ABB RobotStudio station: projekt2.rspag

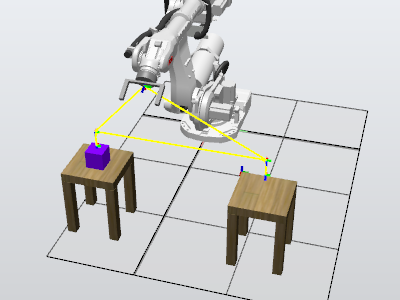
--- station ---
Station Baczyk2 (saved by RobotStudio 24.3.10958.1)
Controller Controller1
  mechanical unit ROB_1: IRB6650S_125_350_MH3_03, 6 joints, base frame (0, 0, 0) mm
Layout (positions relative to the parent item):
  - IRB6650S_125_350_MH3_03 [mechanism, from %ABB.RobotStudio.Models.IRB6650S%\IRB6650S_125_350_MH3_03.rslib] at (0, 0, 0) mm; joint values [0, 0, 0, 0, 0.5236, 0] (rad or m)
  - My_Mechanism [mechanism] at (2365.21, 0, 2010) mm, rotated rx 180 ry 60 rz 180 deg; joint values [0.16, -0.16] (rad or m)
      TCP My_Mechanism_1 at (0, 0, 90) mm
      links: L1, L2, L3
  - Group_2 [graphiccomponentgroup] at (1970.93, 882.73, 0) mm
    - Part_6 [part], size 100 x 100 x 700 mm
    - Part_7 [part], size 100 x 100 x 700 mm
    - Part_8 [part], size 100 x 100 x 700 mm
    - Part_9 [part], size 100 x 100 x 700 mm
    - Part_10 [part], size 600 x 600 x 100 mm
  - Group_3 [graphiccomponentgroup] at (1950.21, -956.94, 0) mm
    - Part_6 [part], size 100 x 100 x 700 mm
    - Part_7 [part], size 100 x 100 x 700 mm
    - Part_8 [part], size 100 x 100 x 700 mm
    - Part_9 [part], size 100 x 100 x 700 mm
    - Part_10 [part], size 600 x 600 x 100 mm
  - LineSensor_2 [smart component, from Components\LineSensor.rslib] at (2444.15, 0, 1965) mm, rotated rx 180 ry 60 rz 180 deg
      properties: Start=[0 0 0]; End=[0 0 0.15]; Length=0.15; Radius=0.01; Tag=(none); SensedPart=(none); SensedPoint=[0 0 0]
    - _sensorPart_ [part], size 20 x 20 x 150 mm
  - Attacher [smart component, from Components\Attacher.rslib]
      properties: Parent=IRB6650S_125_350_MH3_03; Flange=0; Child=(none); Mount=false; Offset=[0 0 0]; Orientation=[0 0 0]
  - Detacher [smart component, from Components\Detacher.rslib]
      properties: Child=(none); KeepPosition=true
  - Part_11 [part] at (2169.73, -741.66, 799.61) mm, size 200 x 200 x 200 mm
  - PoseMover [smart component, from Components\PoseMover.rslib]
      properties: Mechanism=My_Mechanism; Pose=1; Duration=0
  - PoseMover_2 [smart component, from Components\PoseMover.rslib]
      properties: Mechanism=My_Mechanism; Pose=2; Duration=0
  - PoseMover_3 [smart component, from Components\PoseMover.rslib]
      properties: Mechanism=My_Mechanism; Pose=1; Duration=0
Attachment: My_Mechanism is attached to IRB6650S_125_350_MH3_03 / Link6
Attachment: LineSensor_2 is attached to My_Mechanism / L2
EventTableEntry 2426: ActivationMode=2, Cyclic=false, Group=, Trigger=Gripper 2427, Actions=[EventTableActionMechanicalPose 2428], Comment=
EventTableTriggerIO 2427: Operator=0, IOValue=[1], IRC5Controller=? -1, SignalSource=Controller1 2434
EventTableActionMechanicalPose 2428: VirtualSignal=, Mechanism=My_Mechanism 2419, ToPoseName=HomePosition, VirtualSignalValue=[1]
EventTableTriggerIO 2429: Operator=0, IOValue=[0], IRC5Controller=? -1, SignalSource=Controller1 2434
EventTableEntry 2430: ActivationMode=2, Cyclic=false, Group=, Trigger=Gripper 2429, Actions=[EventTableActionMechanicalPose 2431], Comment=
EventTableActionMechanicalPose 2431: VirtualSignal=, Mechanism=My_Mechanism 2419, ToPoseName=SyncPosition, VirtualSignalValue=[1]
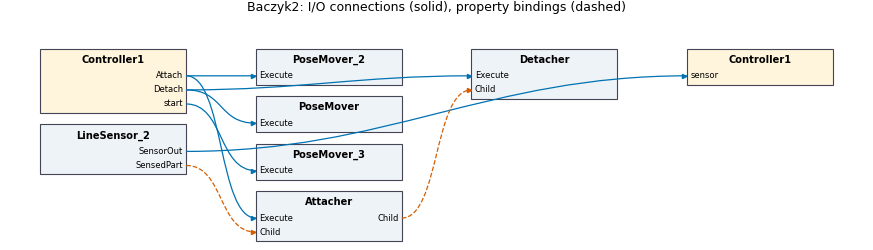
Station logic (signal -> signal, property => property):
  Controller1.Attach -> Attacher.Execute
  Controller1.Detach -> Detacher.Execute
  Controller1.Attach -> PoseMover_2.Execute
  Controller1.Detach -> PoseMover.Execute
  LineSensor_2.SensorOut -> Controller1.sensor
  Controller1.start -> PoseMover_3.Execute
  LineSensor_2.SensedPart => Attacher.Child
  Attacher.Child => Detacher.Child
Targets, tools, work objects and paths stored in the station and not in the controller backup, written as RAPID:
! task T_ROB1
MODULE Module1
  PROC Path_Flow()
    WaitTime 1;
    Set Gripper;
    WaitTime 1;
    Reset Gripper;
    WaitTime 1;
  ENDPROC
ENDMODULE


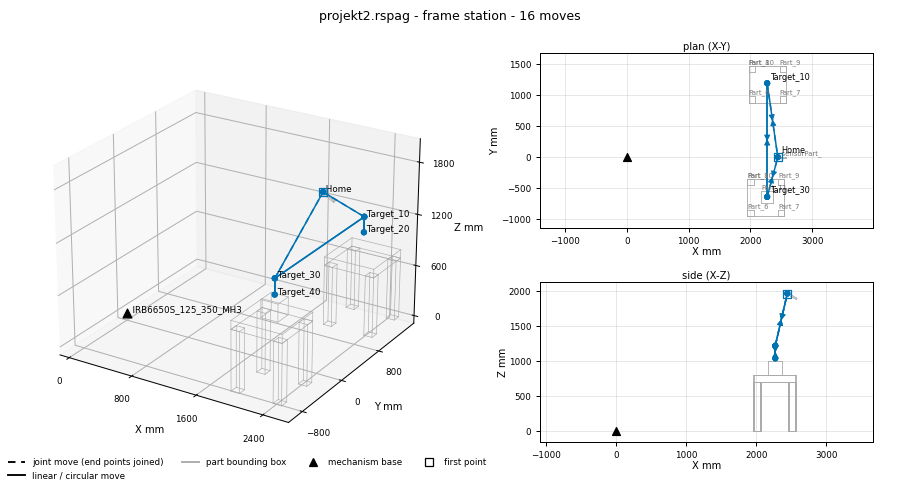
[picture p0: tool path of projekt2.rspag in frame station, 16 of 16 moves have a stored position in this frame; points joined in program order, loops and branches not executed]
--- Controller Data/Controller1/RAPID/TASK1/PROGMOD/CalibData.mod ---
MODULE CalibData
    PERS tooldata My_Mechanism_1:=[TRUE,[[0,0,90],[1,0,0,0]],[1,[0,0,90],[1,0,0,0],0,0,0]];
    TASK PERS wobjdata Workobject_2:=[FALSE,TRUE,"",[[0,0,0],[1,0,0,0]],[[0,0,0],[1,0,0,0]]];
    TASK PERS wobjdata Workobject_3:=[FALSE,TRUE,"",[[1970.926,882.727,800],[1,0,0,0]],[[0,0,0],[1,0,0,0]]];
ENDMODULE

--- Controller Data/Controller1/RAPID/TASK1/PROGMOD/Module1.mod ---
MODULE Module1
    VAR bool value;
        CONST robtarget Home:=[[472.221367097,-882.727,1165],[0.5,0,0.866025404,0],[0,0,0,0],[9E+09,9E+09,9E+09,9E+09,9E+09,9E+09]];
    CONST robtarget Target_10:=[[300.224086373,313.272936929,420.000073654],[-0.000000284,0.000000194,1,-0.000000149],[0,0,0,0],[9E+09,9E+09,9E+09,9E+09,9E+09,9E+09]];
    CONST robtarget Target_20:=[[300.224119695,313.272954476,239.999979637],[-0.000000267,0.000000194,1,-0.00000014],[0,0,0,0],[9E+09,9E+09,9E+09,9E+09,9E+09,9E+09]];
    CONST robtarget Target_30:=[[300.224073663,-1524.727216206,420.000075687],[-0.000000372,0.000000252,1,-0.00000014],[-1,-1,-1,0],[9E+09,9E+09,9E+09,9E+09,9E+09,9E+09]];
    CONST robtarget Target_40:=[[300.224095291,-1524.727007335,240.000010396],[-0.000000007,0,1,0.000000002],[-1,0,-1,0],[9E+09,9E+09,9E+09,9E+09,9E+09,9E+09]];
!***********************************************************
    !
    ! Module:  Module1
    !
    ! Description:
    !   <Insert description here>
    !
    ! Author: Mirgi
    !
    ! Version: 1.0
    !
    !***********************************************************


    !***********************************************************
    !
    ! Procedure main
    !
    !   This is the entry point of your program
    !
    !***********************************************************
    VAR bool detected;
    PROC main()
        Path_10;
    ENDPROC
    PROC Path_10()
        MoveJ Home,v1000,z100,My_Mechanism_1\WObj:=Workobject_3;
        MoveL Target_10,v1000,z100,My_Mechanism_1\WObj:=Workobject_3;
        MoveL Target_20,v1000,fine,My_Mechanism_1\WObj:=Workobject_3;
        IF sensor = 1 THEN
            PulseDO Attach;
            WaitTime 1;
            MoveL Target_10,v1000,z100,My_Mechanism_1\WObj:=Workobject_3;
            MoveL Target_30,v1000,z100,My_Mechanism_1\WObj:=Workobject_3;
            MoveL Target_40,v1000,fine,My_Mechanism_1\WObj:=Workobject_3;
            PulseDO Detach;
            WaitTime 1;
            MoveL Target_30,v1000,z100,My_Mechanism_1\WObj:=Workobject_3;
            MoveJ Home,v1000,z100,My_Mechanism_1\WObj:=Workobject_3;
        ELSE
            MoveJ Home,v1000,z100,My_Mechanism_1\WObj:=Workobject_3;
            MoveL Target_30,v1000,z100,My_Mechanism_1\WObj:=Workobject_3;
            MoveL Target_40,v1000,fine,My_Mechanism_1\WObj:=Workobject_3;
            PulseDO Attach;
            WaitTime 1;
            MoveL Target_30,v1000,z100,My_Mechanism_1\WObj:=Workobject_3;
            MoveL Target_10,v1000,z100,My_Mechanism_1\WObj:=Workobject_3;
            MoveL Target_20,v1000,fine,My_Mechanism_1\WObj:=Workobject_3;
            PulseDO Detach;
            WaitTime 1;
            MoveL Target_10,v1000,z100,My_Mechanism_1\WObj:=Workobject_3;
            MoveJ Home,v1000,z100,My_Mechanism_1\WObj:=Workobject_3;
        ENDIF
    ENDPROC
ENDMODULE

--- Controller Data/Controller1/SYSPAR/EIO.cfg ---
EIO:CFG_1.0:6:1::
#
EIO_SIGNAL:

      -Name "Gripper" -SignalType "DO" -Access "All"

      -Name "Attach" -SignalType "DO"

      -Name "Detach" -SignalType "DO"

      -Name "sensor" -SignalType "DI"

      -Name "start" -SignalType "DO"
